{attribute 'qualified_only'}
{attribute 'to_string'}
TYPE E_Anybus_Media :
(
	eNone				:= 0,	// no sending
	eFirstWater			:= 1,	// pre-rinse, T93 recycle water
	eSoda				:= 2,	// detergent, T92
	eIntermediateWater	:= 3,	// T94 water
	eDisinfection		:= 4,	// T91
	eLastWater			:= 5	// final rinse, T94 water
);
END_TYPE

(* stored: Version 1.1.0.1, ProductVersion 3.1.4026.20
   DUT E_Anybus_Media: Id {c462a162-48be-4fdd-a6ad-b5eaeb29b969} *)
